Fanuc KAREL source: kc00013.KL

-- PROVISIONAL review KL for V770-1; original PC SHA256 f4960ce41c3dbf4a55b554b8eb735d9966502cf1651b66520a231ebe19f7b080
-- Incomplete behavior may be omitted. Consult companion uncertainty JSON. Do not deploy.
PROGRAM KC00013
%NOLOCKGROUP
BEGIN
  -- UNRESOLVED_PC offsets 5-39; opcodes 27,22,22,22,22,22,31
  -- UNRESOLVED_PC offsets 44-48; opcodes 7F
END KC00013
